// TIA Portal V21 export
DATA_BLOCK "Recipe"   // DB30
TITLE = Rezept / Recipe / Recette
{ S7_Optimized_Access := 'TRUE' }
// Werte des Rezepts / Values of the recipe / Valeurs de la recette
   VAR
      target : Int := 500;   // Sollfüllstand in mm / Target level in mm / Niveau de consigne en mm
      hysteresis : Int := 20;   // Hysteresis in mm
   END_VAR
BEGIN
END_DATA_BLOCK
